Fanuc KAREL source: ka00165.KL

-- PROVISIONAL review KL for V770-1; original PC SHA256 ea33a10e65e862164255804c369cf6c2718703b921e74afba3245229eb586ae8
-- Incomplete behavior may be omitted. Consult companion uncertainty JSON. Do not deploy.
PROGRAM KA00165
%NOLOCKGROUP
-- UNRESOLVED_DECL SRC type=002012
-- UNRESOLVED_DECL DST type=002012
BEGIN
  -- UNRESOLVED_PC offsets 5-19; opcodes 22,22,1E
  -- UNRESOLVED_PC offsets 24-28; opcodes 7F
END KA00165
